Fanuc KAREL source: KO00068.KL

PROGRAM KO00068
%NOLOCKGROUP
%ENVIRONMENT MIR
VAR
  P1: XYZWPREXT
  P2: POSITION
  F: BOOLEAN
  OUT: JOINTPOS
BEGIN
  F = TRUE
  OUT = MIRROR(P1, P2, F)
END KO00068
